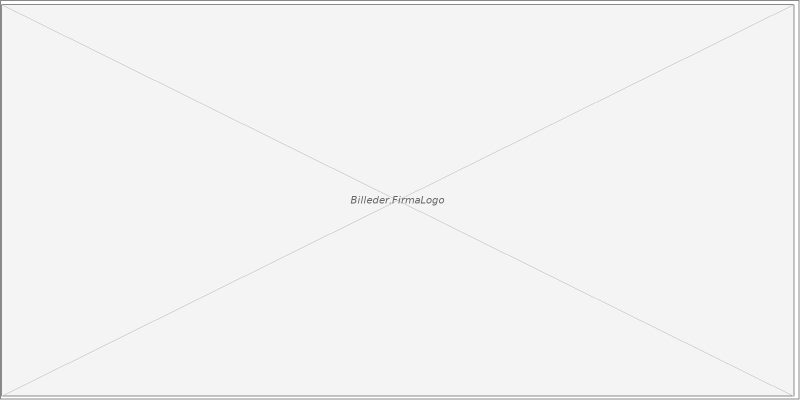
VISUALIZATION Start  // 800x400
    Image (1,4 793x392), image: Billeder.FirmaLogo
END_VISUALIZATION

(* stored: Version 1.1.0.1, ProductVersion 3.1.4024.12
   Visu Start: Id {1ddcc670-8b4f-4c7f-936e-57019fb79669} *)
